(* IEC 61131-3 sources: JingjiangArm/moonboxpro_arm_8.4/Application/Application/任务列表/ExtTask/动作处理/工艺辅助/热风, 2 files *)

(* ---- KS_ReCfgHotBlowerIO.st ---- *)
(*@CES
Name=KS_ReCfgHotBlowerIO
Type=FunctionBlock
TypeGuid=6f9dac99-8de1-4efc-8465-68ac443b7d08
Guid=38ee2e16-ce71-4341-b3d7-8aa23afc131e
HasDeclaration=True
HasImplementation=True
*)
{DECLARATION}
FUNCTION KS_ReCfgHotBlowerIO : BOOL
VAR_INPUT
	i_xInput				: BOOL;(*输入重新分配*)
	i_xOutput				: BOOL;(*输出重新分配*)
	i_xHotBlowerFlag		: BOOL;(*全体热风启动标志*)
	i_iGrpAxisNum_Pu         : INT ;
	i_aiGrpAxisList			: ARRAY [1..MAX_UNIT_NUM] OF INT;(*系的轴列表*)
	i_paxAxisStartEn		: POINTER TO ARRAY [1..MAX_UNIT_NUM] OF BOOL;(*轴启动使能|有效后按钮开关才能起作用*)
	i_paxStartKnob			: POINTER TO ARRAY [1..MAX_UNIT_NUM] OF BOOL;(*全体启动,每个轴旋钮输入*)
	i_paxStartOrStopBtn		: POINTER TO ARRAY [1..MAX_UNIT_NUM] OF BOOL;(*单轴的启动停止按钮*)
	i_paxNeedStop			: POINTER TO ARRAY [1..MAX_UNIT_NUM] OF BOOL;(*单轴需要停止标志*)
	i_paxAxisStarted		: POINTER TO ARRAY [1..MAX_UNIT_NUM] OF BOOL;(*单个轴的启动输出标志|实际处于启动状态，
																			可以根据i_paxNeedStop这个变量控制实际输出*)
	i_byHotBlowerStopDelayTime: BYTE;(*热风延时关闭时间|S*)
	i_patAxisDelayTimeSa	: POINTER TO ARRAY [1..MAX_UNIT_NUM] OF TIME;(*延时开始时间|用于和当前时间对比检查是否到时间*)
	i_pxFlag_AxisStopping   : POINTER TO BOOL;(*热风停止中|至少一个轴*)
	i_axHotBlower :ARRAY [1..MAX_UNIT_NUM] OF BOOL;
	i_axHotBlower_Button:ARRAY [1..MAX_UNIT_NUM] OF BOOL;
	i_axHotBlower_Err:ARRAY [1..MAX_UNIT_NUM] OF BOOL;
	i_axLamp_Heating:ARRAY [1..MAX_UNIT_NUM] OF BOOL;
	i_paxRel_HotBlower:POINTER TO ARRAY [1..MAX_UNIT_NUM] OF BOOL;
	i_paxLamp_HotBlower:POINTER TO ARRAY [1..MAX_UNIT_NUM] OF BOOL;
	i_paxLamp_AllHotBlower:POINTER TO ARRAY [1..MAX_UNIT_NUM] OF BOOL;
	i_pxLamp_AllHotBlower		:POINTER TO BOOL;
END_VAR
VAR
	iUnitId: INT;
	iN: INT;
	xAxisStartEn: BOOL;
	xNeedStop: BOOL;
	tTimeCur: TIME;
	xAxisSts: BOOL;
	axAxisStoping		:  ARRAY [1..MAX_UNIT_NUM] OF BOOL;(*轴热风停止中|用于加热时延时关闭*)
	xFlag_AxisStopping	: BOOL;
END_VAR

{IMPLEMENTATION}
IF i_paxAxisStartEn<>0 AND
	i_paxStartKnob<>0 AND
	i_paxNeedStop<>0 AND
 	i_paxStartOrStopBtn<>0 AND
	i_paxAxisStarted<>0 AND
	i_pxFlag_AxisStopping<>0 AND
	i_patAxisDelayTimeSa<>0 THEN
	tTimeCur:=TIME();
	IF i_xInput THEN
		FOR iN:=1 TO MAX_UNIT_NUM  BY 1 DO
			i_paxStartKnob^[iN]:=FALSE;
			i_paxStartOrStopBtn^[iN]:=FALSE;
			i_paxNeedStop^[iN]:=FALSE;
			i_paxAxisStartEn^[iN]:=FALSE;
		END_FOR

		FOR iN:=1 TO i_iGrpAxisNum_Pu  BY 1 DO
			iUnitId:=i_aiGrpAxisList[iN];
			IF iUnitId>0 AND iUnitId<= MAX_UNIT_NUM THEN
				i_paxStartKnob^[iUnitId]:=i_axHotBlower[iUnitId];
				i_paxStartOrStopBtn^[iUnitId]:=i_axHotBlower_Button[iUnitId];
				xNeedStop:=i_axHotBlower_Err[iUnitId];
				i_paxNeedStop^[iUnitId]:=xNeedStop;

				xAxisStartEn:=TRUE;
				i_paxAxisStartEn^[iUnitId]:=xAxisStartEn;
			END_IF
		END_FOR
	ELSIF i_xOutput THEN
		FOR iN:=1 TO i_iGrpAxisNum_Pu  BY 1 DO
			iUnitId:=i_aiGrpAxisList[iN];
			IF iUnitId>0 AND iUnitId <= MAX_UNIT_NUM THEN(*输出循环到收牵，这样热风输出灯就可以配到收牵上了|2020.1.9.094955*)
				IF i_paxAxisStarted^[iUnitId] THEN(*如果打开的话|我们直接输出临时变量*)
					xAxisSts:=TRUE;
				ELSE(*关闭时  保持之前状态*)
					IF i_byHotBlowerStopDelayTime=0 THEN(*延时=0的时候直接关闭*)
						xAxisSts:=FALSE;
					ELSE
						xAxisSts:=i_paxRel_HotBlower^[iUnitId];
					END_IF
					IF xAxisSts THEN(**)
						axAxisStoping[iUnitId]:=TRUE;(*停止过程中*)
					END_IF
				END_IF

				(*2021.7.27.115739  增加了加热打开时 热风延时关闭|*)
				IF i_axLamp_Heating[iUnitId] THEN(*处于加热过程中|保留当前时间*)
					i_patAxisDelayTimeSa^[iUnitId]:=tTimeCur;
				ELSE(*加热关闭了|统计关闭时间-*)
					IF tTimeCur-i_patAxisDelayTimeSa^[iUnitId]>=WORD_TO_TIME(BYTE_TO_WORD(i_byHotBlowerStopDelayTime)*1000) THEN(*时间到了|如果需要关闭，可正常关闭*)
						IF NOT i_paxAxisStarted^[iUnitId] THEN(*热风关闭的时候*)
							xAxisSts:=FALSE;
							axAxisStoping[iUnitId]:=FALSE;
						END_IF
					ELSE;
					END_IF
				END_IF

				IF axAxisStoping[iUnitId] THEN(*有一个轴停止中|*)
					xFlag_AxisStopping:=TRUE;
				END_IF

				i_paxLamp_HotBlower^[iUnitId]:=(*i_paxAxisStarted^[iUnitId]*)xAxisSts;
				i_paxRel_HotBlower^[iUnitId]:=(*i_paxAxisStarted^[iUnitId]*)xAxisSts;
(*				i_pastStIOMap_AxisExtra^[iUnitId].o_xLamp_AllHotBlower:=i_xHotBlowerFlag OR xFlag_AxisStopping;*)
			END_IF
		END_FOR

		FOR iN:=1 TO i_iGrpAxisNum_Pu + 2  BY 1 DO
			(*输出到牵引，*)
			IF  iN >=  i_iGrpAxisNum_Pu THEN
				i_pxLamp_AllHotBlower^ :=  i_xHotBlowerFlag OR xFlag_AxisStopping;;
			ELSE
				iUnitId:=i_aiGrpAxisList[iN];
				IF iUnitId>0 AND iUnitId <= MAX_UNIT_NUM THEN(*输出循环到收牵，这样热风输出灯就可以配到收牵上了|2020.1.9.094955*)
					i_paxLamp_AllHotBlower^[iUnitId]:=i_xHotBlowerFlag OR xFlag_AxisStopping;
				END_IF
			END_IF
		END_FOR
		i_pxFlag_AxisStopping^:=xFlag_AxisStopping;
	END_IF
END_IF

(* ---- KS_FB_GrpAirHotCtrl.st ---- *)
(*@CES
Name=KS_FB_GrpAirHotCtrl
Type=FunctionBlock
TypeGuid=6f9dac99-8de1-4efc-8465-68ac443b7d08
Guid=1e8a028d-d061-44b5-a7fa-8fcf2eecc751
HasDeclaration=True
HasImplementation=True
*)
{DECLARATION}
FUNCTION_BLOCK KS_FB_GrpAirHotCtrl
(*2020.10.13.133218 重新处理热风功能|Liu.yt*)
(*2024.7.1.165726 循环索引增加到了i_iGrpAxisTotalNum*)
VAR_INPUT
	i_xEn: BOOL;
	i_iGrpAxisNum_Pu: INT; (*色组轴数*)
	i_iAxisId_If  : INT ;
	i_iAxisId_Of : INT;
	i_iGrpId	:INT ;
	i_aiGrpAxisList: ARRAY [1..MAX_UNIT_NUM] OF INT; (*系的轴列表*)
	i_pstStEvtReq:POINTER TO StEvtReq;
	i_xHotBlowerByKnob:BOOL;(*单轴启动根据旋钮开关标志|用于全体开关控制启动的逻辑|无则不输入*)
	i_xAirExhaustFinishFlag:BOOL;(*排风完成标志*)
	i_xAirExhaustLimit:BOOL;(*排风限制热风*)
	i_xStopHotBlowerWhenEstop:BOOL;(*急停停止热风标志|有效了和急停关联，无效则不影响*)
	i_iCycleTime_Plc:INT;(*2024.01.22.142933+*)

	i_pstStSysParam  : POINTER TO StSysParam   ; (*系统参数*)
	i_PastStIOMap_Axis_Extra_FE:  POINTER TO ARRAY [1..MAX_UNIT_NUM] OF StIOMap_Axis_Extra_FE  ;
	i_pastStIOMap_Main_FE	: POINTER TO ARRAY [1..4] OF StIOMap_Main_FE;(*轴io数据区域|*)
END_VAR
VAR_OUTPUT
	o_xEno: BOOL;
	o_iErNo: INT;(*0成功\-1参数无效|*)
	o_xHotBlowerFlag:BOOL;(*热风启动标志*)
	o_xFlag_HotBlowerStopping:BOOL;(*热风停止中*)
	o_axHotBlowerEn: ARRAY [1..MAX_UNIT_NUM] OF BOOL;(*热风启动标志|停止时和实际输出存在不一致*)
	o_axHotBlowerEn_Act: ARRAY [1..MAX_UNIT_NUM] OF BOOL;(*热风启动标志和读取实际反馈*)
END_VAR
VAR

	fbKS_FB_HotBlowerSys: KS_FB_BlowerFunction;
	axAxisStartKnob: ARRAY [1..MAX_UNIT_NUM] OF BOOL;
	axStartOrStopBtn: ARRAY [1..MAX_UNIT_NUM] OF BOOL;
	axNeedStop: ARRAY [1..MAX_UNIT_NUM] OF BOOL;
	axAxisStartEn: ARRAY [1..MAX_UNIT_NUM] OF BOOL;
	xHotBlowerEn: BOOL;
	iStartedSum: INT;(*启动的轴数*)
	iN: INT;
	iUnitId:INT;

	atHotBlowerDelayTimeSa: ARRAY [1..MAX_UNIT_NUM] OF TIME;
	byHotBlowerStopDelayTime_In : BYTE ;
	iDelayMsec_HeatBlower_In : INT  ;
	xFlag_Estop_In: BOOL;
	axHotBlower_In :ARRAY [1..MAX_UNIT_NUM] OF BOOL;
	axHotBlower_Button_In :ARRAY [1..MAX_UNIT_NUM] OF BOOL;
	axHotBlower_Err_In :ARRAY [1..MAX_UNIT_NUM] OF BOOL;
	axLamp_Heating_In :ARRAY [1..MAX_UNIT_NUM] OF BOOL;
	axHotBlower_Opened_Act_In :ARRAY [1..MAX_UNIT_NUM] OF BOOL;

	axRel_HotBlower_Out : ARRAY [1..MAX_UNIT_NUM] OF BOOL;
	axLamp_HotBlower_Out: ARRAY [1..MAX_UNIT_NUM] OF BOOL;
	axLamp_AllHotBlower_Out:ARRAY [1..MAX_UNIT_NUM] OF BOOL;

	xLamp_AllHotBlower_Out: BOOL;

	pstStUnitParam_Save: POINTER TO  StUnitParam_Save;
	pstStIOMap_Axis_Extra_FE:  POINTER TO  StIOMap_Axis_Extra_FE  ;
END_VAR
{IMPLEMENTATION}
Action_Input();

Action_ActCtl() ;

Action_Output();
